// TIA Portal V20 export
ORGANIZATION_BLOCK "T2_Ciclo"   // OB125, LAD, ProgramCycle
TITLE = T2_Ciclo
{ S7_Optimized_Access := 'TRUE' }
AUTHOR : IA
FAMILY : PRUEBA
VERSION : 0.1
// Prueba IA 2: llama a todas las pruebas base en cada ciclo
// stored: AutoNumber false, IsIECCheckEnabled false, SetENOAutomatically false
   VAR_INPUT
      Initial_Call : Bool;
      Remanence : Bool;
   END_VAR
BEGIN

REGION Network 1: Contador de vida
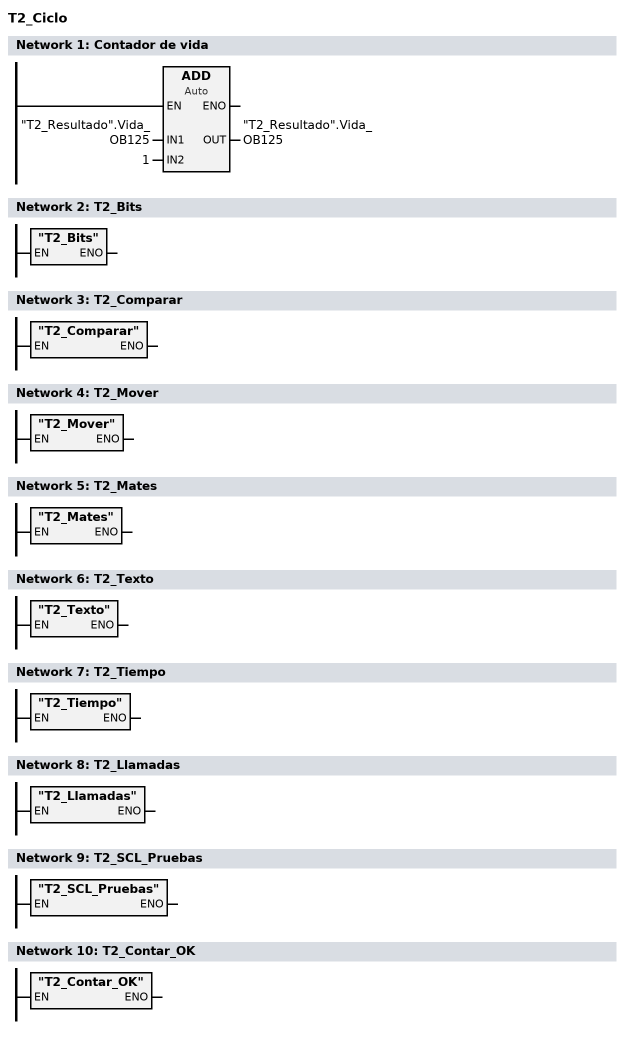
   RUNG wire#powerrail
      Add(in1 := "T2_Resultado".Vida_OB125, in2 := 1, out => "T2_Resultado".Vida_OB125)
   END_RUNG
   // the same network as SCL:
   "T2_Resultado".Vida_OB125 := "T2_Resultado".Vida_OB125 + 1;
END_REGION

REGION Network 2: T2_Bits
   RUNG wire#powerrail
      "T2_Bits"()
   END_RUNG
   // the same network as SCL:
   "T2_Bits"();
END_REGION

REGION Network 3: T2_Comparar
   RUNG wire#powerrail
      "T2_Comparar"()
   END_RUNG
   // the same network as SCL:
   "T2_Comparar"();
END_REGION

REGION Network 4: T2_Mover
   RUNG wire#powerrail
      "T2_Mover"()
   END_RUNG
   // the same network as SCL:
   "T2_Mover"();
END_REGION

REGION Network 5: T2_Mates
   RUNG wire#powerrail
      "T2_Mates"()
   END_RUNG
   // the same network as SCL:
   "T2_Mates"();
END_REGION

REGION Network 6: T2_Texto
   RUNG wire#powerrail
      "T2_Texto"()
   END_RUNG
   // the same network as SCL:
   "T2_Texto"();
END_REGION

REGION Network 7: T2_Tiempo
   RUNG wire#powerrail
      "T2_Tiempo"()
   END_RUNG
   // the same network as SCL:
   "T2_Tiempo"();
END_REGION

REGION Network 8: T2_Llamadas
   RUNG wire#powerrail
      "T2_Llamadas"()
   END_RUNG
   // the same network as SCL:
   "T2_Llamadas"();
END_REGION

REGION Network 9: T2_SCL_Pruebas
   RUNG wire#powerrail
      "T2_SCL_Pruebas"()
   END_RUNG
   // the same network as SCL:
   "T2_SCL_Pruebas"();
END_REGION

REGION Network 10: T2_Contar_OK
   RUNG wire#powerrail
      "T2_Contar_OK"()
   END_RUNG
   // the same network as SCL:
   "T2_Contar_OK"();
END_REGION
END_ORGANIZATION_BLOCK
